(* IEC 61131-3 sources: llm-plc-st-eval/data/definitivo/gemini-3.1-pro-preview/I7/few_shot, 3 files *)

(* ---- ejec_1.st ---- *)
FUNCTION_BLOCK FB_Duplex
VAR_INPUT
    demanda : BOOL; (* Senal de arranque del grupo *)
    falla1 : BOOL;  (* Falla de la bomba 1 *)
    falla2 : BOOL;  (* Falla de la bomba 2 *)
END_VAR
VAR_OUTPUT
    bomba1 : BOOL;   (* Comando de la bomba 1 *)
    bomba2 : BOOL;   (* Comando de la bomba 2 *)
    almFalla : BOOL; (* Alarma de falla en bomba principal *)
END_VAR
VAR
    rTrigDemanda : R_TRIG; (* Detector de flanco de subida de la demanda *)
    turnoBomba2 : BOOL := TRUE; (* Inicia en TRUE para que la primera demanda asigne el turno a la bomba 1 *)
END_VAR

(* Deteccion de nueva demanda para alternar el turno *)
rTrigDemanda(CLK := demanda);
IF rTrigDemanda.Q THEN
    turnoBomba2 := NOT turnoBomba2;
END_IF;

(* Logica de control de bombas y alarmas *)
IF demanda THEN
    IF NOT turnoBomba2 THEN
        (* Bomba 1 es la principal *)
        bomba1 := NOT falla1;
        bomba2 := falla1 AND NOT falla2;
        almFalla := falla1;
    ELSE
        (* Bomba 2 es la principal *)
        bomba2 := NOT falla2;
        bomba1 := falla2 AND NOT falla1;
        almFalla := falla2;
    END_IF;
ELSE
    (* Sin demanda, ambas bombas y la alarma se apagan *)
    bomba1 := FALSE;
    bomba2 := FALSE;
    almFalla := FALSE;
END_IF;
END_FUNCTION_BLOCK

(* ---- ejec_2.st ---- *)
FUNCTION_BLOCK FB_Duplex
VAR_INPUT
    demanda : BOOL; (* Señal de demanda de bombeo *)
    falla1  : BOOL; (* Falla de la bomba 1 *)
    falla2  : BOOL; (* Falla de la bomba 2 *)
END_VAR
VAR_OUTPUT
    bomba1   : BOOL; (* Comando de arranque bomba 1 *)
    bomba2   : BOOL; (* Comando de arranque bomba 2 *)
    almFalla : BOOL; (* Alarma de falla en bomba principal *)
END_VAR
VAR
    rTrigDemanda : R_TRIG; (* Detector de flanco de subida de la demanda *)
    turnoBomba1  : BOOL := FALSE; (* Alternancia, inicia en FALSE para que el primer cambio sea a TRUE *)
END_VAR

(* Alternar la bomba principal en cada nueva demanda (transicion de FALSE a TRUE) *)
rTrigDemanda(CLK := demanda);
IF rTrigDemanda.Q THEN
    turnoBomba1 := NOT turnoBomba1;
END_IF;

(* Control de bombas y alarma segun la demanda y el turno *)
IF demanda THEN
    IF turnoBomba1 THEN
        (* Bomba 1 es principal, Bomba 2 es respaldo *)
        bomba1 := NOT falla1;
        bomba2 := falla1 AND NOT falla2;
        almFalla := falla1;
    ELSE
        (* Bomba 2 es principal, Bomba 1 es respaldo *)
        bomba2 := NOT falla2;
        bomba1 := falla2 AND NOT falla1;
        almFalla := falla2;
    END_IF;
ELSE
    (* Sin demanda, ambas bombas y la alarma se apagan *)
    bomba1 := FALSE;
    bomba2 := FALSE;
    almFalla := FALSE;
END_IF;
END_FUNCTION_BLOCK

(* ---- ejec_3.st ---- *)
FUNCTION_BLOCK FB_Duplex
VAR_INPUT
    demanda : BOOL; (* Peticion de arranque *)
    falla1 : BOOL;  (* Falla de la bomba 1 *)
    falla2 : BOOL;  (* Falla de la bomba 2 *)
END_VAR
VAR_OUTPUT
    bomba1 : BOOL;   (* Comando de arranque bomba 1 *)
    bomba2 : BOOL;   (* Comando de arranque bomba 2 *)
    almFalla : BOOL; (* Alarma de falla en la bomba principal *)
END_VAR
VAR
    flancoDemanda : R_TRIG; (* Detector de flanco de subida *)
    bomba1Principal : BOOL := FALSE; (* Alternancia: inicia en FALSE para que el primer pulso lo haga TRUE *)
END_VAR

(* Deteccion de nueva demanda para alternar el rol de bomba principal *)
flancoDemanda(CLK := demanda);
IF flancoDemanda.Q THEN
    bomba1Principal := NOT bomba1Principal;
END_IF;

(* La bomba 1 arranca si hay demanda, no tiene falla, y es la principal o la bomba 2 (principal) fallo *)
bomba1 := demanda AND NOT falla1 AND (bomba1Principal OR falla2);

(* La bomba 2 arranca si hay demanda, no tiene falla, y es la principal o la bomba 1 (principal) fallo *)
bomba2 := demanda AND NOT falla2 AND (NOT bomba1Principal OR falla1);

(* La alarma se activa solo si hay demanda y la bomba que tiene el rol principal presenta falla *)
almFalla := demanda AND ((bomba1Principal AND falla1) OR (NOT bomba1Principal AND falla2));
END_FUNCTION_BLOCK
